// TIA Portal V21 export
// export: Created 2026-11-10T07:35:06.0726591Z, ExportSetting WithDefaults, DisplayName Totally Integrated Automation Portal, DisplayVersion V21 Update 3, DisplayName STEP 7 Professional, DisplayVersion V21 Update 3, DisplayName STEP 7 Safety, DisplayVersion V21, DisplayName Tech WebApplication, DisplayVersion V21, DisplayName WinCC Basic/Comfort/Advanced, DisplayVersion V21 Update 3, DisplayName WinCC Unified, DisplayVersion V21 Update 3
FUNCTION_BLOCK "FB_Lad_ex048"   // FB93, LAD
{ S7_Optimized_Access := 'TRUE' }
VERSION : 0.1
// stored: AutoNumber true, IsIECCheckEnabled false, IsRetainMemResEnabled false, MemoryReserve 100, SetENOAutomatically false, UDAEnableTagReadback false
   VAR_INPUT
      v_id : HW_SUBMODULE;
   END_VAR
   VAR_OUTPUT
      v_status : DWord;
   END_VAR
   VAR_IN_OUT
      v_outputs : Array[0..99] of Byte;
   END_VAR
   VAR
      inst { S7_SetPoint := 'True'} : SETIO;
   END_VAR
BEGIN

REGION Network 1: SETIO - Write all outputs of a submodule
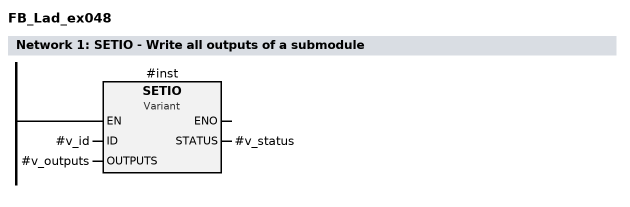
   RUNG wire#powerrail
      { S7_Templates := "[card := 0, ptr_type := Variant, id_type := HW_SUBMODULE]" } #inst.SETIO(ID := #v_id, STATUS => #v_status, OUTPUTS := #v_outputs)
   END_RUNG
   // the same network as SCL:
   #inst(ID := #v_id, OUTPUTS := #v_outputs, STATUS => #v_status);   // SETIO
END_REGION
END_FUNCTION_BLOCK
